(* IEC 61131-3 sources: TetherPLC/tests/tempctrl/cases, 21 files *)

(* ---- t13_handoff.st ---- *)
// t13_handoff.st — the WebUI autotune handoff shape, runtime-verified.
// Mirrors what fbd-lower's expand_st_blocks generates for an inline
// `st` block: VAR_IN_OUT pins aliasing tuner/controller FB instances,
// VAR_OUTPUT live mirrors, and a one-shot APPLY strobe copying gains
// into the controller's input members (CTL.K1 := TUNE.K1 …).
// Same model params as t06 → K1≈6.188 K2≈1.089 Ki≈0.671.
FUNCTION_BLOCK FB_TuneHandoff
VAR_INPUT
    APPLY : BOOL;
    RESET : BOOL;
END_VAR
VAR_OUTPUT
    lqr_k1 : LREAL;
    lqr_k2 : LREAL;
    lqr_ki : LREAL;
    lqr_done : BOOL;
END_VAR
VAR_IN_OUT
    TUNE : FB_AtcLqrTune;
    CTL : FB_AtcLqr;
END_VAR
VAR
    applied : BOOL;
END_VAR
    lqr_k1 := TUNE.K1;
    lqr_k2 := TUNE.K2;
    lqr_ki := TUNE.Ki;
    lqr_done := TUNE.Done;
    IF APPLY AND NOT applied THEN
        CTL.K1 := TUNE.K1;
        CTL.K2 := TUNE.K2;
        CTL.Ki := TUNE.Ki;
        applied := TRUE;
    END_IF;
    IF RESET THEN applied := FALSE; END_IF;
END_FUNCTION_BLOCK

PROGRAM T13
VAR
    flags AT %QB0 : BYTE;
    m : FB_AtcModel2s;
    t : FB_AtcLqrTune;
    c : FB_AtcLqr;
    ho : FB_TuneHandoff;
END_VAR
    m(Execute := TRUE, K := 1.0, Tau := 20.0, Theta := 0.0,
      TauH := 5.0, Ts := 0.5);
    t(Execute := TRUE, A11 := m.A11, A12 := m.A12,
      A21 := m.A21, A22 := m.A22, B1 := m.B1, B2 := m.B2,
      Q1 := 1.0, Q2 := 0.1, Qi := 0.5, R := 1.0, Ts := 0.5,
      MaxIter := 0, Tol := 0.0);
    // K1/K2/Ki intentionally omitted — the handoff owns them; binding
    // them here would clobber the tuned gains every scan (same reason
    // applyTunerToPou strips those params from the controller block).
    c(Execute := FALSE, Setpoint := 0.0, Actual := 0.0,
      X2 := 0.0,
      Nref := 0.0, FFwd := 0.0, OutMin := -100.0, OutMax := 100.0,
      RateLim := 0.0, ManEn := FALSE, ManOut := 0.0,
      CycleTime := 0.1, Reset := FALSE);
    ho(TUNE := t, CTL := c, APPLY := TRUE, RESET := FALSE);
    flags := 0;
    IF t.Done AND t.Conv THEN flags := flags + 1; END_IF;
    IF ABS(ho.lqr_k1 - t.K1) < 0.001 THEN flags := flags + 2; END_IF;
    IF c.K1 > 6.0 AND c.K1 < 6.4 THEN flags := flags + 4; END_IF;
    IF c.K2 > 1.0 AND c.K2 < 1.2 THEN flags := flags + 8; END_IF;
    IF c.Ki > 0.6 AND c.Ki < 0.75 THEN flags := flags + 16; END_IF;
END_PROGRAM

(* ---- t01_math.st ---- *)
// t01_math.st — math function conformance: exp/ln/sqrt/pow against
// known values; flags bit i set when the check passes.
PROGRAM T01
VAR
    flags AT %QB0 : BYTE;
    e1 AT %QD8 : LREAL;
    l1 AT %QD16 : LREAL;
    s1 AT %QD24 : LREAL;
    p1 AT %QD32 : LREAL;
    l2 AT %QD40 : LREAL;
    s2 AT %QD48 : LREAL;
END_VAR
    e1 := F_AtcExp(1.0);          // e = 2.718281828...
    l1 := F_AtcLn(F_AtcExp(3.7)); // = 3.7
    s1 := F_AtcSqrt(2.0);         // 1.41421356...
    p1 := F_AtcPow(2.0, 10.0);    // 1024
    l2 := F_AtcLn(100.0);         // 4.605170186
    s2 := F_AtcSqrt(0.001);       // 0.031622776
    flags := 0;
    IF e1 > 2.718281 AND e1 < 2.718282 THEN flags := flags + 1; END_IF;
    IF l1 > 3.6999 AND l1 < 3.7001 THEN flags := flags + 2; END_IF;
    IF s1 > 1.414213 AND s1 < 1.414214 THEN flags := flags + 4; END_IF;
    IF p1 > 1023.999 AND p1 < 1024.001 THEN flags := flags + 8; END_IF;
    IF l2 > 4.605169 AND l2 < 4.605171 THEN flags := flags + 16; END_IF;
    IF s2 > 0.031622 AND s2 < 0.031624 THEN flags := flags + 32; END_IF;
END_PROGRAM

(* ---- t02_pid.st ---- *)
// t02_pid.st — FB_AtcPid closed loop on a simulated first-order
// plant (K=2 deg/%, Tau=10 s, Ts=0.5 s): PI must pull PV from 20 to
// SP=80 and hold it there. flags: b0 PV in band, b1 output in range,
// b2 Done, b3 no error, b4 anti-windup: output never exceeded 100.
PROGRAM T02
VAR
    flags AT %QB0 : BYTE;
    c : FB_AtcPid;
    pv : LREAL;
    u AT %QD8 : LREAL;
    pvO AT %QD16 : LREAL;
    satHist : LREAL;
END_VAR
    c(Execute := TRUE, Setpoint := 80.0, Actual := pv,
      Kp := 3.0, Tn := 8.0, Tv := 0.0, TfD := 0.0,
      B := 1.0, C := 0.0, FFwd := 0.0,
      OutMin := 0.0, OutMax := 100.0, RateLim := 0.0,
      Deadband := 0.0, HoldI := FALSE, TrackEn := FALSE,
      TrackVal := 0.0, ManEn := FALSE, ManOut := 0.0,
      CycleTime := 0.5, Reset := FALSE);
    u := c.Out;
    IF u > 100.01 OR u < -0.01 THEN
        satHist := 1.0;
    END_IF;
    // plant lag (start PV at 20 deg)
    pv := pv + (2.0 * u - pv) * (0.5 / (10.0 + 0.5));
    pvO := pv;
    flags := 0;
    IF pv > 78.5 AND pv < 82.5 THEN flags := flags + 1; END_IF;
    IF u >= 0.0 AND u <= 100.0 THEN flags := flags + 2; END_IF;
    IF c.Done THEN flags := flags + 4; END_IF;
    IF NOT c.Err THEN flags := flags + 8; END_IF;
    IF satHist = 0.0 THEN flags := flags + 16; END_IF;
END_PROGRAM

(* ---- t03_relay.st ---- *)
// t03_relay.st — FB_AtcRelayTune on a simulated first-order plant
// (K=1, Tau=10 s, Ts=0.5 s): relay hysteresis 2 deg around SP=50,
// MeanOut=50, amp=20. Must finish with Done, plausible Ku/Tu, and
// ZN-classic gains Kp=0.6Ku Tn=0.5Tu Tv=0.125Tu.
// flags: b0 Done, b1 Ku in [4,20], b2 Tu in [4,60], b3 Kp>0,
//        b4 Tn=0.5*Tu, b5 Tv=0.125*Tu, b6 Busy went low, b7 no Err.
PROGRAM T03
VAR
    flags AT %QB0 : BYTE;
    c : FB_AtcRelayTune;
    pv : LREAL;
    u AT %QD8 : LREAL;
    kuO AT %QD16 : LREAL;
    tuO AT %QD24 : LREAL;
END_VAR
    c(Execute := TRUE, Setpoint := 50.0, Actual := pv,
      RelayAmp := 20.0, MeanOut := 50.0, Hyst := 2.0,
      OutMin := 0.0, OutMax := 100.0, TuneRule := 0,
      MinCyc := 3, CycleTime := 0.5,
      Abort := FALSE, Reset := FALSE);
    u := c.Out;
    pv := pv + (1.0 * u - pv) * (0.5 / (10.0 + 0.5));
    kuO := c.Ku;
    tuO := c.Tu;
    flags := 0;
    IF c.Done THEN flags := flags + 1; END_IF;
    IF c.Ku > 4.0 AND c.Ku < 30.0 THEN flags := flags + 2; END_IF;
    IF c.Tu > 4.0 AND c.Tu < 40.0 THEN flags := flags + 4; END_IF;
    IF c.Kp > 0.0 THEN flags := flags + 8; END_IF;
    IF ABS(c.Tn - 0.5 * c.Tu) < 0.01 THEN flags := flags + 16; END_IF;
    IF ABS(c.Tv - 0.125 * c.Tu) < 0.01 THEN flags := flags + 32; END_IF;
    IF NOT c.Busy THEN flags := flags + 64; END_IF;
    IF NOT c.Err THEN flags := flags + 128; END_IF;
END_PROGRAM

(* ---- t04_stepid.st ---- *)
// t04_stepid.st — FB_AtcStepIdent on a simulated FOPDT plant:
// K=2 deg/%, Tau=20 s, true delay 7.5 s (15-scan shift at Ts=0.5),
// step U0=10 -> U1=40. Expect K~2, Tau~20, Theta~7.5+lag bias.
// flags: b0 Done, b1 |K-2|<0.15, b2 14<Tau<28, b3 4<Theta<14,
//        b4 Busy low, b5 no Err, b6 PvFinal ~ K*U1 = 80.
PROGRAM T04
VAR
    flags AT %QB0 : BYTE;
    id : FB_AtcStepIdent;
    pv : LREAL;
    dl : ARRAY[0..15] OF LREAL;
    i : DINT;
    u AT %QD8 : LREAL;
    kO AT %QD16 : LREAL;
    tauO AT %QD24 : LREAL;
    thO AT %QD32 : LREAL;
END_VAR
    id(Execute := TRUE, Actual := pv, U0 := 10.0, U1 := 40.0,
       SettleT := 120.0, TolBand := 0.05, SettleN := 8,
       MaxTime := 600.0, StoreEvery := 4, CycleTime := 0.5,
       Reset := FALSE);
    u := id.Out;
    // plant: 7.5 s transport delay + 20 s lag, gain 2
    pv := pv + (2.0 * dl[15] - pv) * (0.5 / (20.0 + 0.5));
    FOR i := 0 TO 14 DO
        dl[15 - i] := dl[14 - i];
    END_FOR;
    dl[0] := u;
    kO := id.K;
    tauO := id.Tau;
    thO := id.Theta;
    flags := 0;
    IF id.Done THEN flags := flags + 1; END_IF;
    IF id.K > 1.85 AND id.K < 2.15 THEN flags := flags + 2; END_IF;
    IF id.Tau > 14.0 AND id.Tau < 28.0 THEN flags := flags + 4; END_IF;
    IF id.Theta > 4.0 AND id.Theta < 14.0 THEN flags := flags + 8; END_IF;
    IF NOT id.Busy THEN flags := flags + 16; END_IF;
    IF NOT id.Err THEN flags := flags + 32; END_IF;
    IF id.PvFinal > 75.0 AND id.PvFinal < 85.0 THEN
        flags := flags + 64;
    END_IF;
END_PROGRAM

(* ---- t05_rules.st ---- *)
// t05_rules.st — FB_AtcTuneRules on a known FOPDT model
// (K=2, Tau=20, Theta=5). Rule 0 IMC lambda=max(1.25,4)=4:
//   Kp=(20+2.5)/(2*(4+2.5))=1.7308 Tn=22.5 Tv=100/45=2.2222
// Rule 1 SIMC lambda=5: Kp=20/(2*10)=1.0 Tn=min(20,40)=20 Tv=0
// flags: b0 IMC done, b1..3 IMC values, b4 SIMC done, b5 SIMC Kp,
//        b6 ZN done, b7 ZN Kp = 1.2*20/(2*5) = 2.4
PROGRAM T05
VAR
    flags AT %QB0 : BYTE;
    r0 : FB_AtcTuneRules;
    r1 : FB_AtcTuneRules;
    r2 : FB_AtcTuneRules;
    kp0 AT %QD8 : LREAL;
    kp1 AT %QD16 : LREAL;
END_VAR
    r0(Execute := TRUE, K := 2.0, Tau := 20.0, Theta := 5.0,
       Rule := 0, Lambda := 0.0);
    r1(Execute := TRUE, K := 2.0, Tau := 20.0, Theta := 5.0,
       Rule := 1, Lambda := 0.0);
    r2(Execute := TRUE, K := 2.0, Tau := 20.0, Theta := 5.0,
       Rule := 2, Lambda := 0.0);
    kp0 := r0.Kp;
    kp1 := r1.Kp;
    flags := 0;
    IF r0.Done THEN flags := flags + 1; END_IF;
    IF r0.Kp > 1.70 AND r0.Kp < 1.76 THEN flags := flags + 2; END_IF;
    IF r0.Tn > 22.4 AND r0.Tn < 22.6 THEN flags := flags + 4; END_IF;
    IF r0.Tv > 2.2 AND r0.Tv < 2.3 THEN flags := flags + 8; END_IF;
    IF r1.Done THEN flags := flags + 16; END_IF;
    IF r1.Kp > 0.99 AND r1.Kp < 1.01 THEN flags := flags + 32; END_IF;
    IF r2.Done THEN flags := flags + 64; END_IF;
    IF r2.Kp > 2.39 AND r2.Kp < 2.41 THEN flags := flags + 128; END_IF;
END_PROGRAM

(* ---- t06_tuners.st ---- *)
// t06_tuners.st — solvers vs reference values.
// Model from FB_AtcModel2s for K=1 Tau=20 TauH=5 Theta=0 Ts=0.5:
//   a1=e^(-0.025)=0.9753099 a2=e^(-0.1)=0.9048374
//   A=[[.9753,.0247],[0,.9048]] B=[0,0.09516]
// FB_AtcLqrTune Q=diag(1,0.1,0.5) R=1 ->
//   ref (scipy DARE, -Ts aug): K1=6.1884 K2=1.0892 Ki=0.6712
// FB_AtcKalmanTune Q=diag(.01,.01) R=1 -> L1=0.0777 L2=0.00609
// flags: b0/b4 done+conv, b1..3 K in range, b5..6 L in range,
//        b7 model outputs in range
PROGRAM T06
VAR
    flags AT %QB0 : BYTE;
    m : FB_AtcModel2s;
    t : FB_AtcLqrTune;
    kf : FB_AtcKalmanTune;
    k1 AT %QD8 : LREAL;
    k2 AT %QD16 : LREAL;
    ki AT %QD24 : LREAL;
    l1 AT %QD32 : LREAL;
END_VAR
    m(Execute := TRUE, K := 1.0, Tau := 20.0, Theta := 0.0,
      TauH := 5.0, Ts := 0.5);
    t(Execute := TRUE, A11 := m.A11, A12 := m.A12,
      A21 := m.A21, A22 := m.A22, B1 := m.B1, B2 := m.B2,
      Q1 := 1.0, Q2 := 0.1, Qi := 0.5, R := 1.0, Ts := 0.5,
      MaxIter := 0, Tol := 0.0);
    kf(Execute := TRUE, A11 := m.A11, A12 := m.A12,
       A21 := m.A21, A22 := m.A22,
       Q1 := 0.01, Q2 := 0.01, R := 1.0,
       MaxIter := 0, Tol := 0.0);
    k1 := t.K1;
    k2 := t.K2;
    ki := t.Ki;
    l1 := kf.L1;
    flags := 0;
    IF m.Done THEN flags := flags + 1; END_IF;
    IF t.K1 > 6.0 AND t.K1 < 6.4 THEN flags := flags + 2; END_IF;
    IF t.K2 > 1.0 AND t.K2 < 1.2 THEN flags := flags + 4; END_IF;
    IF t.Ki > 0.6 AND t.Ki < 0.75 THEN flags := flags + 8; END_IF;
    IF t.Done AND t.Conv THEN flags := flags + 16; END_IF;
    IF kf.Done AND kf.Conv THEN flags := flags + 32; END_IF;
    IF kf.L1 > 0.07 AND kf.L1 < 0.09 THEN flags := flags + 64; END_IF;
    IF kf.L2 > 0.004 AND kf.L2 < 0.008 THEN flags := flags + 128; END_IF;
END_PROGRAM

(* ---- t07_lqr.st ---- *)
// t07_lqr.st — FB_AtcLqr closed loop on the discrete 2-state sim it
// was tuned for (same A/B as t06). K1=6.1884 K2=1.0892 Ki=0.6712,
// Nref=0 (integral does the tracking). SP=80, x1 starts 0.
// flags: b0 x1 in band, b1 Out in range, b2 Done, b3 no Err,
//        b4 xi finite.
PROGRAM T07
VAR
    flags AT %QB0 : BYTE;
    c : FB_AtcLqr;
    x1 : LREAL;
    x2 : LREAL;
    u AT %QD8 : LREAL;
END_VAR
    c(Execute := TRUE, Setpoint := 80.0, Actual := x1, X2 := x2,
      K1 := 6.1884, K2 := 1.0892, Ki := 0.6712,
      Nref := 0.0, FFwd := 0.0,
      OutMin := 0.0, OutMax := 100.0, RateLim := 0.0,
      ManEn := FALSE, ManOut := 0.0,
      CycleTime := 0.5, Reset := FALSE);
    u := c.Out;
    // plant (discrete, Ts=0.5): x1+ = a1 x1 + (1-a1) x2
    //                         x2+ = a2 x2 + K(1-a2) u
    x1 := 0.9753099 * x1 + 0.0246901 * x2;
    x2 := 0.9048374 * x2 + 0.0951626 * u;
    flags := 0;
    IF x1 > 79.0 AND x1 < 81.0 THEN flags := flags + 1; END_IF;
    IF u >= -0.01 AND u <= 100.01 THEN flags := flags + 2; END_IF;
    IF c.Done THEN flags := flags + 4; END_IF;
    IF NOT c.Err THEN flags := flags + 8; END_IF;
    IF c.Xi > -1.0e6 AND c.Xi < 1.0e6 THEN flags := flags + 16; END_IF;
END_PROGRAM

(* ---- t08_lqg.st ---- *)
// t08_lqg.st — FB_AtcLqg closed loop: same plant as t07 but PV is
// corrupted by a deterministic +/- noise square wave (amplitude 0.5);
// the Kalman filter (L1=0.0777 L2=0.00609) must still track.
// flags: b0 x1 plant state in band, b1 estimated X1 near PV mean,
//        b2 Out bounded, b3 Done, b4 no Err, b5 X2 estimate finite.
PROGRAM T08
VAR
    flags AT %QB0 : BYTE;
    c : FB_AtcLqg;
    x1 : LREAL;
    x2 : LREAL;
    nz : LREAL;
    ymeas : LREAL;
    u AT %QD8 : LREAL;
    xe AT %QD16 : LREAL;
END_VAR
    // deterministic measurement noise: +-0.5 alternating every 7 scans
    nz := nz + 0.5;
    IF nz >= 7.0 THEN nz := -7.0; END_IF;
    ymeas := x1 + nz / 7.0 * 0.5 - 0.25;
    c(Execute := TRUE, Setpoint := 80.0, Actual := ymeas,
      A11 := 0.9753099, A12 := 0.0246901,
      A21 := 0.0, A22 := 0.9048374,
      B1 := 0.0, B2 := 0.0951626,
      L1 := 0.0777, L2 := 0.00609,
      K1 := 6.1884, K2 := 1.0892, Ki := 0.6712,
      Nref := 0.0, FFwd := 0.0,
      OutMin := 0.0, OutMax := 100.0,
      ManEn := FALSE, ManOut := 0.0,
      CycleTime := 0.5, Reset := FALSE);
    u := c.Out;
    x1 := 0.9753099 * x1 + 0.0246901 * x2;
    x2 := 0.9048374 * x2 + 0.0951626 * u;
    xe := c.X1;
    flags := 0;
    IF x1 > 78.0 AND x1 < 82.0 THEN flags := flags + 1; END_IF;
    IF c.X1 > 78.0 AND c.X1 < 82.0 THEN flags := flags + 2; END_IF;
    IF u >= -0.01 AND u <= 100.01 THEN flags := flags + 4; END_IF;
    IF c.Done THEN flags := flags + 8; END_IF;
    IF NOT c.Err THEN flags := flags + 16; END_IF;
    IF c.X2 > -1.0e6 AND c.X2 < 1.0e6 THEN flags := flags + 32; END_IF;
END_PROGRAM

(* ---- t09_profile.st ---- *)
// t09_profile.st — FB_AtcProfile exercising all segment kinds:
//   SEG1 RAMP  -> 100 at 4 deg/s   (PV start 20 -> ~20 s)
//   SEG2 DWELL    100 for 30 s, guaranteed-soak band 2.0
//   SEG3 RAMPT -> 60 in 40 s
//   SEG4 STEP  -> 60 (jump, EV pulse)
//   SEG5 LOOP  -> seg 2, x1 (dwell+rampt run twice)
//   SEG6 END
// Simulated PV lags SP at 10 s. flags: b0 ran to END (Done),
// b1 SP hit 100, b2 SegIdx visited 2, b3 EV word seen (seg2 EV=2),
// b4 guaranteed soak stretched dwell (dwell seg took > 30 s while
// PV lagging outside band... here PV tracks so gsoak rarely bites;
// instead check dwell SegIdx stayed for >= 30 s), b5 loop ran twice
// (saw SegIdx=2 twice => SegIdx reached 4 then 2 again), b6 SP
// finished at 60 (RAMPT target of second pass), b7 no Err.
PROGRAM T09
VAR
    flags AT %QB0 : BYTE;
    prof : FB_AtcProfile;
    pv : LREAL;
    sp AT %QD8 : LREAL;
    segO AT %QD16 : DINT;
    run : BOOL;
    cnt : DINT;
    sawDwell : DINT;
    dwellStart : LREAL;
    dwellLong : BOOL;
    sawSeg4 : BOOL;
    sawLoop : BOOL;
END_VAR
    // ---- segment table (member-wise writes; aggregates can't bind)
    IF cnt = 0 THEN
        prof.SEG[1].KIND := 2;  // RAMP
        prof.SEG[1].TGT := 100.0;
        prof.SEG[1].P1 := 4.0;
        prof.SEG[1].EV := 1;
        prof.SEG[2].KIND := 1;  // DWELL
        prof.SEG[2].TGT := 100.0;
        prof.SEG[2].P1 := 30.0;
        prof.SEG[2].P2 := 2.0;
        prof.SEG[2].EV := 2;
        prof.SEG[3].KIND := 3;  // RAMPT
        prof.SEG[3].TGT := 60.0;
        prof.SEG[3].P1 := 40.0;
        prof.SEG[3].EV := 4;
        prof.SEG[4].KIND := 4;  // STEP
        prof.SEG[4].TGT := 60.0;
        prof.SEG[4].EV := 8;
        prof.SEG[5].KIND := 5;  // LOOP -> seg 2, 1 extra pass
        prof.SEG[5].TGT := 2.0;
        prof.SEG[5].P1 := 1.0;
        prof.SEG[6].KIND := 0;  // END
    END_IF;
    cnt := cnt + 1;
    IF cnt = 2 THEN
        pv := 20.0;   // PV-start point
        run := TRUE;
    END_IF;
    prof(NUM_SEG := 6, RUN := run, HOLD := FALSE, RESET := FALSE,
         PvStart := TRUE, PV := pv, CycleTime := 0.5);
    run := FALSE;
    // simulated PV follows SP (1st-order, 10 s lag)
    pv := pv + (prof.SP - pv) * (0.5 / (10.0 + 0.5));
    sp := prof.SP;
    segO := prof.SegIdx;
    // book-keeping for checks
    IF prof.SegIdx = 2 THEN
        sawDwell := sawDwell + 1;
        IF sawDwell = 1 THEN dwellStart := prof.SegTime; END_IF;
    END_IF;
    IF prof.SegIdx = 2 AND prof.SegTime >= 29.5 THEN
        dwellLong := TRUE;
    END_IF;
    IF prof.SegIdx = 4 THEN sawSeg4 := TRUE; END_IF;
    IF sawSeg4 AND prof.SegIdx = 2 THEN sawLoop := TRUE; END_IF;
    flags := 0;
    IF prof.Done THEN flags := flags + 1; END_IF;
    IF sawDwell >= 2 THEN flags := flags + 2; END_IF;
    IF dwellLong THEN flags := flags + 4; END_IF;
    IF sawSeg4 THEN flags := flags + 8; END_IF;
    IF sawLoop THEN flags := flags + 16; END_IF;
    IF prof.SP > 59.0 AND prof.SP < 61.0 THEN
        flags := flags + 32;
    END_IF;
    IF NOT prof.Err THEN flags := flags + 64; END_IF;
    // extra: the EV word of the END segment is 0; while busy it was
    // nonzero at least once — sawLoop covers seg-2 revisit.
    IF prof.Busy OR prof.Done THEN flags := flags + 128; END_IF;
END_PROGRAM

(* ---- t10_cascade.st ---- *)
// t10_cascade.st — FB_AtcCascadePid: outer product loop (slow, Tau=30)
// drives inner heater loop (fast, Tau=2) setpoint range 20..150;
// inner drives duty 0..100 with gain 1.5 deg/%.
// flags: b0 product PV within band, b1 inner SP clamped to range,
//        b2 Out in range, b3 Done, b4 no Err.
PROGRAM T10
VAR
    flags AT %QB0 : BYTE;
    c : FB_AtcCascadePid;
    pvO : LREAL;
    pvI : LREAL;
    u AT %QD8 : LREAL;
    ispO AT %QD16 : LREAL;
    badIsp : BOOL;
END_VAR
    c(Execute := TRUE, Setpoint := 80.0,
      PvOuter := pvO, PvInner := pvI,
      KpO := 2.0, TnO := 40.0, TvO := 0.0,
      KpI := 4.0, TnI := 4.0, TvI := 0.0,
      InnerSpMin := 20.0, InnerSpMax := 150.0,
      OutMin := 0.0, OutMax := 100.0,
      ManEn := FALSE, ManOut := 0.0,
      CycleTime := 0.5, Reset := FALSE);
    u := c.Out;
    ispO := c.InnerSp;
    IF c.InnerSp < 19.99 OR c.InnerSp > 150.01 THEN
        badIsp := TRUE;
    END_IF;
    // plants: heater lag Tau=2 gain 1.5; product follows heater Tau=30
    pvI := pvI + (1.5 * u - pvI) * (0.5 / (2.0 + 0.5));
    pvO := pvO + (pvI - pvO) * (0.5 / (30.0 + 0.5));
    flags := 0;
    IF pvO > 77.0 AND pvO < 83.0 THEN flags := flags + 1; END_IF;
    IF NOT badIsp THEN flags := flags + 2; END_IF;
    IF u >= -0.01 AND u <= 100.01 THEN flags := flags + 4; END_IF;
    IF c.Done THEN flags := flags + 8; END_IF;
    IF pvI > 0.0 AND pvI <= 150.01 THEN flags := flags + 16; END_IF;
END_PROGRAM

(* ---- t11_smith.st ---- *)
// t11_smith.st — FB_AtcSmith on a dead-time plant:
// K=1 deg/%, Tau=8 s, delay=7.5 s (15 scans); model identical.
// The dead-time compensation must hold SP=60 without oscillation.
// flags: b0 PV in band, b1 Out in range, b2 Done, b3 no Err,
//        b4 model delay state nonzero.
PROGRAM T11
VAR
    flags AT %QB0 : BYTE;
    c : FB_AtcSmith;
    pv : LREAL;
    dl : ARRAY[0..15] OF LREAL;
    i : DINT;
    u AT %QD8 : LREAL;
END_VAR
    c(Execute := TRUE, Setpoint := 60.0, Actual := pv,
      Kp := 0.6, Tn := 10.0, Tv := 0.0,
      ModelK := 1.0, ModelT := 8.0, ModelDt := 7.5,
      OutMin := 0.0, OutMax := 100.0,
      ManEn := FALSE, ManOut := 0.0,
      CycleTime := 0.5, Reset := FALSE);
    u := c.Out;
    // plant: 15-scan delay + 8 s lag, gain 1
    pv := pv + (1.0 * dl[15] - pv) * (0.5 / (8.0 + 0.5));
    FOR i := 0 TO 14 DO
        dl[15 - i] := dl[14 - i];
    END_FOR;
    dl[0] := u;
    flags := 0;
    IF pv > 58.0 AND pv < 62.5 THEN flags := flags + 1; END_IF;
    IF u >= -0.01 AND u <= 100.01 THEN flags := flags + 2; END_IF;
    IF c.Done THEN flags := flags + 4; END_IF;
    IF NOT c.Err THEN flags := flags + 8; END_IF;
    IF c.E > -100.0 AND c.E < 100.0 THEN flags := flags + 16; END_IF;
END_PROGRAM

(* ---- t12_util.st ---- *)
// t12_util.st — signal helpers: FB_AtcPt1, FB_AtcRateLim,
// FB_AtcPwm, FB_AtcHeatCool.
// flags: b0 Pt1 near input after 10*timeconst scans,
//        b1 RateLim respected (|dOut| <= Rate*Ts + eps),
//        b2 Pwm duty ~50% over a period (count on-scans),
//        b3 HeatCool splits (U=-40 -> Cool=40-DeadZone),
//        b4 all Done.
PROGRAM T12
VAR
    flags AT %QB0 : BYTE;
    f1 : FB_AtcPt1;
    rl : FB_AtcRateLim;
    pw : FB_AtcPwm;
    hc : FB_AtcHeatCool;
    cnt : DINT;
    onCnt : DINT;
    pv : LREAL;
    rlPrev : LREAL;
    rlOk : BOOL;
    rlIn : LREAL;
END_VAR
    cnt := cnt + 1;
    // Pt1: step 0->50 at scan 1, Tf=4s
    f1(Execute := TRUE, In := 50.0, Tf := 4.0,
       CycleTime := 0.5, Reset := FALSE);
    pv := f1.Out;
    // RateLim: square wave input +-20, Rate=10/s -> |dOut| <= 5/scan
    IF cnt >= 100 THEN rlIn := -20.0; ELSE rlIn := 20.0; END_IF;
    rl(Execute := TRUE, In := rlIn, Rate := 10.0,
       CycleTime := 0.5, Reset := FALSE);
    IF cnt > 1 THEN
        IF rl.Out - rlPrev > 5.001 OR rl.Out - rlPrev < -5.001 THEN
            rlOk := TRUE;
        END_IF;
    END_IF;
    rlPrev := rl.Out;
    // Pwm: Duty=50, Period=4s (8 scans) — count on-scans over 8 scans
    pw(Execute := TRUE, Duty := 50.0, Period := 4.0, MinOn := 0.0,
       CycleTime := 0.5, Reset := FALSE);
    IF cnt > 190 AND cnt <= 198 THEN
        IF pw.Q THEN onCnt := onCnt + 1; END_IF;
    END_IF;
    // HeatCool: U=-40, dz=2 -> Cool=38*1=38
    hc(Execute := TRUE, U := -40.0, DeadZone := 2.0, CoolGain := 1.0);
    flags := 0;
    IF pv > 48.0 AND pv <= 50.0 THEN flags := flags + 1; END_IF;
    IF NOT rlOk THEN flags := flags + 2; END_IF;
    IF onCnt >= 3 AND onCnt <= 5 THEN flags := flags + 4; END_IF;
    IF hc.Cool > 37.9 AND hc.Cool < 38.1 AND hc.Heat = 0.0 THEN
        flags := flags + 8;
    END_IF;
    IF f1.Done AND rl.Done AND pw.Done AND hc.Done THEN
        flags := flags + 16;
    END_IF;
END_PROGRAM

(* ---- t14_aiscale.st ---- *)
// t14_aiscale.st — FB_AtcAiScale / FB_AtcAoScale: raw int16 channel
// counts <-> engineering units, incl. PT1 filtering and int16
// saturation. Sticky check bits compose into flags %QB0 at the end
// of every scan (idempotent): b0 ai linear exact, b1 ai filtered
// converging, b2 ao roundtrip, b3 ao saturates high, b4 ao
// saturates low -> expect 0x1f.
PROGRAM T14
VAR
    flags AT %QB0 : BYTE;
    ok0, ok1, ok2, ok3, ok4 : BOOL;
    ai : FB_AtcAiScale;
    aoRT : FB_AtcAoScale;
    aoHi : FB_AtcAoScale;
    aoLo : FB_AtcAoScale;
    aiF : FB_AtcAiScale;
    raw : INT;               // analog input channel counts (EL3104-style)
    rawF : INT;              // second channel for the filter test
    counts : INT;            // analog output channel counts (EL4104-style)
    ct : LREAL;
    n : DINT;
END_VAR
    ct := 0.1;
    n := n + 1;

    // ---- AI: EU = Raw*Scale + Offset, no filter
    IF n = 1 THEN raw := 16384; END_IF;
    ai(Execute := TRUE, Raw := raw, Scale := 0.5, Offset := 10.0,
       FiltT := 0.0, CycleTime := ct, Reset := FALSE);
    // 16384 * 0.5 + 10 = 8202
    IF ai.Done AND ai.Out > 8201.9 AND ai.Out < 8202.1 THEN
        ok0 := TRUE;
    END_IF;

    // ---- AI filtered: FiltT=1 s, ct=0.1 -> alpha = 0.1/1.1
    // step rawF 0 -> 1100 counts at n=20; rawf approaches 1100
    IF n = 20 THEN rawF := 1100; END_IF;
    aiF(Execute := TRUE, Raw := rawF, Scale := 1.0, Offset := 0.0,
        FiltT := 1.0, CycleTime := ct, Reset := FALSE);
    // after ~40 filtered steps rawf ~= 1100*(1-(1-alpha)^40) ~ 1080
    IF n >= 40 AND aiF.RawF > 1000.0 AND aiF.RawF < 1100.0 THEN
        ok1 := TRUE;
    END_IF;

    // ---- AO: counts = (In - Offset)/Scale -> int16
    aoRT(Execute := TRUE, In := 8202.0, Scale := 0.5, Offset := 10.0,
         CycleTime := ct, Reset := FALSE);
    IF aoRT.Done AND aoRT.Counts = 16384 AND NOT aoRT.OutBad THEN
        ok2 := TRUE;
    END_IF;

    // ---- AO saturation: way over range -> rail + OutBad
    aoHi(Execute := TRUE, In := 40000.0, Scale := 0.5, Offset := 10.0,
         CycleTime := ct, Reset := FALSE);
    IF aoHi.Done AND aoHi.Counts >= 32767 AND aoHi.OutBad THEN
        ok3 := TRUE;
    END_IF;
    aoLo(Execute := TRUE, In := -40000.0, Scale := 0.5, Offset := 10.0,
         CycleTime := ct, Reset := FALSE);
    IF aoLo.Done AND aoLo.Counts <= -32768 AND aoLo.OutBad THEN
        ok4 := TRUE;
    END_IF;

    flags := 0;
    IF ok0 THEN flags := flags + 1; END_IF;
    IF ok1 THEN flags := flags + 2; END_IF;
    IF ok2 THEN flags := flags + 4; END_IF;
    IF ok3 THEN flags := flags + 8; END_IF;
    IF ok4 THEN flags := flags + 16; END_IF;

    // settle: feed AO counts back to image for observability
    counts := aoRT.Counts;
END_PROGRAM

(* ---- t15_lethality.st ---- *)
// t15_lethality.st — FB_AtcLethality: Tref=70, Z=10, F0Target=1.0 min,
// Temp=90 -> rate=10^2/60=1.667 F0/min, +0.1667/scan. InProduct from
// n=1: F0 hits 1.0 at n=6 (Done). ExitProduct pulse n=4 catches
// acc=0.667<target -> Divert. SensorOK drops n=20 -> Frozen latches;
// ExitProduct n=25 diverts on freeze. Reset n=30 clears acc but the
// same scan re-accumulates, so F0=0.167 at n=30.
// Sticky bits -> flags %QB0: expect 0x3f.
PROGRAM T15
VAR
    flags AT %QB0 : BYTE;
    ok0, ok1, ok2, ok3, ok4, ok5 : BOOL;
    le : FB_AtcLethality;
    n : DINT;
    sok, ex : BOOL;
END_VAR
    n := n + 1;
    sok := NOT (n >= 20 AND n <= 29);
    ex := (n = 4) OR (n = 25);
    le(Temp := 90.0, InProduct := TRUE, SensorOK := sok,
       ExitProduct := ex, Tref := 70.0, Z := 10.0,
       F0Target := 1.0, CycleTime := 0.1,
       Reset := (n = 30));
    IF n = 5 AND le.F0 > 0.5 AND le.F0 < 0.9 THEN ok0 := TRUE; END_IF;
    IF n >= 7 AND n < 15 AND le.Done THEN ok1 := TRUE; END_IF;
    IF n = 4 AND le.Divert THEN ok2 := TRUE; END_IF;
    IF n >= 21 AND n <= 24 AND le.Frozen THEN ok3 := TRUE; END_IF;
    IF n = 25 AND le.Divert THEN ok4 := TRUE; END_IF;
    IF n = 30 AND le.F0 < 0.3 THEN ok5 := TRUE; END_IF;
    flags := 0;
    IF ok0 THEN flags := flags + 1; END_IF;
    IF ok1 THEN flags := flags + 2; END_IF;
    IF ok2 THEN flags := flags + 4; END_IF;
    IF ok3 THEN flags := flags + 8; END_IF;
    IF ok4 THEN flags := flags + 16; END_IF;
    IF ok5 THEN flags := flags + 32; END_IF;
END_PROGRAM

(* ---- t16_heatch.st ---- *)
// t16_heatch.st — FB_AtcHeaterChannel: auto PWM phase, interlock
// inhibit, manual select, and duty clamp. n drives the phases:
//   1-10   auto MV=50%, Period=1s, CycleTime=0.1 -> Q toggles
//   11-20  InterlockOK=FALSE -> Q=FALSE, InterlockBad=TRUE
//   21-30  Auto=FALSE, ManualMV=25 -> DutyApplied=25
//   31-35  MV=150 -> DutyApplied clamped to 100
//   36-45  Execute=FALSE -> Q=FALSE, InterlockBad=FALSE
// Sticky bits -> flags %QB0: expect 0x1f.
PROGRAM T16
VAR
    flags AT %QB0 : BYTE;
    ok0, ok1, ok2, ok3, ok4 : BOOL;
    hc : FB_AtcHeaterChannel;
    n : DINT;
    sawQ : BOOL;
END_VAR
    n := n + 1;
    hc.Execute := n <= 35;
    hc.Enable := TRUE;
    hc.Auto := NOT (n >= 21 AND n <= 30);
    hc.MV := 50.0;
    IF n >= 31 THEN hc.MV := 150.0; END_IF;
    hc.ManualMV := 25.0;
    hc.InterlockOK := NOT (n >= 11 AND n <= 20);
    hc.Period := 1.0;
    hc.MinOn := 0.0;
    hc.CycleTime := 0.1;
    hc();
    IF hc.Q THEN sawQ := TRUE; END_IF;
    ok0 := sawQ;
    IF (n = 15) AND hc.InterlockBad AND NOT hc.Q THEN
        ok1 := TRUE;
    END_IF;
    IF (n = 25) AND (hc.DutyApplied = 25.0) THEN
        ok2 := TRUE;
    END_IF;
    IF (n = 33) AND (hc.DutyApplied = 100.0) THEN
        ok3 := TRUE;
    END_IF;
    IF (n = 40) AND NOT hc.Q AND NOT hc.InterlockBad THEN
        ok4 := TRUE;
    END_IF;
    flags := 0;
    IF ok0 THEN flags := flags + 1; END_IF;
    IF ok1 THEN flags := flags + 2; END_IF;
    IF ok2 THEN flags := flags + 4; END_IF;
    IF ok3 THEN flags := flags + 8; END_IF;
    IF ok4 THEN flags := flags + 16; END_IF;
END_PROGRAM

(* ---- t17_plant.st ---- *)
// t17_plant.st — FB_AtcPlant: FOPDT+deadtime plant simulator.
// Phase 1 (cycles 0..39, U=50 open loop): PV must stay near Pv0
// early (Theta=2 s dead time at 0.5 s scan) then rise toward
// K*U = 100.  Phase 2 (cycles 40+, PI control SP=80): PV settles
// in band.  flags: b0 settled, b1 no err, b2 plant Done,
// b3 output in range, b4 heated above 60, b5 dead time held PV<30
// at cycle 4.
PROGRAM T17
VAR
    flags AT %QB0 : BYTE;
    plant : FB_AtcPlant;
    pid : FB_AtcPid;
    cyc : DINT;
    u : LREAL;
    pvEarly : LREAL;
    maxPv : LREAL;
    closed : BOOL;
END_VAR
    cyc := cyc + 1;
    closed := cyc > 40;
    IF closed THEN
        pid(Execute := TRUE, Setpoint := 80.0, Actual := plant.PV,
            Kp := 3.0, Tn := 8.0, Tv := 0.0, TfD := 0.0,
            B := 1.0, C := 0.0, FFwd := 0.0,
            OutMin := 0.0, OutMax := 100.0, RateLim := 0.0,
            Deadband := 0.0, HoldI := FALSE, TrackEn := FALSE,
            TrackVal := 0.0, ManEn := FALSE, ManOut := 0.0,
            CycleTime := 0.5, Reset := FALSE);
        u := pid.Out;
    ELSE
        u := 50.0;
    END_IF;
    plant(Execute := TRUE, U := u, K := 2.0, Tau1 := 10.0,
          Tau2 := 0.0, Theta := 2.0, Pv0 := 20.0, DistU := 0.0,
          Taamb := 20.0, TauAmb := 0.0, NoiseAmp := 0.0,
          CycleTime := 0.5, Reset := cyc = 1);
    IF cyc = 4 THEN pvEarly := plant.PV; END_IF;
    IF plant.PV > maxPv THEN maxPv := plant.PV; END_IF;
    flags := 0;
    IF closed AND plant.PV > 74.0 AND plant.PV < 86.0 THEN
        flags := flags + 1;
    END_IF;
    IF NOT plant.Err AND NOT pid.Err THEN flags := flags + 2; END_IF;
    IF plant.Done THEN flags := flags + 4; END_IF;
    IF u >= 0.0 AND u <= 100.0 THEN flags := flags + 8; END_IF;
    IF maxPv > 60.0 THEN flags := flags + 16; END_IF;
    IF pvEarly > 0.0 AND pvEarly < 30.0 THEN flags := flags + 32; END_IF;
END_PROGRAM

(* ---- t18_trend.st ---- *)
// t18_trend.st — FB_AtcTrend ring-buffer capture.  Depth=64,
// Value=cycle index, Reset on cycle 1 (records start cycle 2),
// trigger at cycle 20 -> ring pos 18, PostN=4.  72 writes total:
// Wr=70, Full wraps at write 64.
// flags: b0 Done, b1 Full, b2 TrigIdx=18, b3 Buf[TrigIdx]=20
// (trigger sample, not yet overwritten), b4 Count>=40, b5 Wr=72 mod 64 = 8.
PROGRAM T18
VAR
    flags AT %QB0 : BYTE;
    tr : FB_AtcTrend;
    cyc : DINT;
END_VAR
    cyc := cyc + 1;
    tr(Execute := TRUE, CycleTime := 0.1,
       Value := DINT_TO_LREAL(cyc), Depth := 64, PostN := 4,
       Arm := TRUE, Trig := cyc = 20, Reset := cyc = 1);
    flags := 0;
    IF tr.Done THEN flags := flags + 1; END_IF;
    IF tr.Full THEN flags := flags + 2; END_IF;
    IF tr.TrigIdx = 18 THEN flags := flags + 4; END_IF;
    IF tr.TrigIdx >= 0 THEN
        IF tr.Buf[tr.TrigIdx] = 20.0 THEN flags := flags + 8; END_IF;
    END_IF;
    IF tr.Count >= 40 THEN flags := flags + 16; END_IF;
    IF tr.Wr = 8 THEN flags := flags + 32; END_IF;
END_PROGRAM

(* ---- t19_gsched.st ---- *)
// t19_gsched.st — FB_AtcGainSchedule breakpoint interpolation.
// Tables configured once as instance members (array call-args do not
// bind in the MIR), then X varies per call.  X=[0,50,100],
// Kp=[1,2,4], Tn=[10,20,40], Tv=[0,1,2].
// flags: b0 X=0  -> Kp=1 Seg=1 Frac=0
//        b1 X=50 -> Kp=2 Seg=1 Frac=1
//        b2 X=25 -> Kp=1.5 Tn=15 Tv=0.5 Frac=0.5
//        b3 X=75 -> Kp=3 Tn=30 Tv=1.5 Seg=2 Frac=0.5
//        b4 X=-10-> Kp=1 (clamp low)
//        b5 X=200-> Kp=4 (clamp high)
//        b6 dup-X table -> Err
//        b7 X=100-> Kp=4 Seg=2 Frac=1
PROGRAM T19
VAR
    flags AT %QB0 : BYTE;
    gs : FB_AtcGainSchedule;
    gb : FB_AtcGainSchedule;
    cyc : DINT;
END_VAR
    cyc := cyc + 1;
    IF cyc = 1 THEN
        gs.TableX[1] := 0.0;   gs.TableX[2] := 50.0;  gs.TableX[3] := 100.0;
        gs.TableKp[1] := 1.0;  gs.TableKp[2] := 2.0;  gs.TableKp[3] := 4.0;
        gs.TableTn[1] := 10.0; gs.TableTn[2] := 20.0; gs.TableTn[3] := 40.0;
        gs.TableTv[1] := 0.0;  gs.TableTv[2] := 1.0;  gs.TableTv[3] := 2.0;
        gb.TableX := gs.TableX;
        gb.TableKp := gs.TableKp;
        gb.TableTn := gs.TableTn;
        gb.TableTv := gs.TableTv;
        gb.TableX[2] := gb.TableX[1];   // duplicate X -> must flag Err
    END_IF;
    IF cyc >= 2 THEN
        flags := 0;
        gs(Execute := TRUE, X := 0.0, NPts := 3);
        IF gs.Kp = 1.0 AND gs.Seg = 1 AND gs.Frac = 0.0 THEN
            flags := flags + 1;
        END_IF;
        gs(Execute := TRUE, X := 50.0, NPts := 3);
        IF gs.Kp = 2.0 AND gs.Seg = 1 AND gs.Frac = 1.0 THEN
            flags := flags + 2;
        END_IF;
        gs(Execute := TRUE, X := 25.0, NPts := 3);
        IF gs.Kp = 1.5 AND gs.Tn = 15.0 AND gs.Tv = 0.5
           AND gs.Frac = 0.5 THEN
            flags := flags + 4;
        END_IF;
        gs(Execute := TRUE, X := 75.0, NPts := 3);
        IF gs.Kp = 3.0 AND gs.Tn = 30.0 AND gs.Tv = 1.5
           AND gs.Seg = 2 AND gs.Frac = 0.5 THEN
            flags := flags + 8;
        END_IF;
        gs(Execute := TRUE, X := -10.0, NPts := 3);
        IF gs.Kp = 1.0 THEN flags := flags + 16; END_IF;
        gs(Execute := TRUE, X := 200.0, NPts := 3);
        IF gs.Kp = 4.0 THEN flags := flags + 32; END_IF;
        gb(Execute := TRUE, X := 10.0, NPts := 3);
        IF gb.Err THEN flags := flags + 64; END_IF;
        gs(Execute := TRUE, X := 100.0, NPts := 3);
        IF gs.Kp = 4.0 AND gs.Seg = 2 AND gs.Frac = 1.0 THEN
            flags := flags + 128;
        END_IF;
    END_IF;
END_PROGRAM

(* ---- t20_autotune.st ---- *)
// t20_autotune.st — FB_AtcAutoTune end-to-end: relay tune on
// FB_AtcPlant (K=1, Tau=10, Theta=1) drives the plant to a limit
// cycle, gains latch, PID takes over bumplessly via TrackEn.
// flags: b0 at.Done seen, b1 gains sane (Kp>0 Tn>0 Tv>=0 Ku>0 Tu>0),
//        b2 PID settled |PV-50|<10 at end, b3 no Err ever,
//        b4 handoff continuity |dOut|<8 at Done scan,
//        b5 Cycles>=2, b6 PidTrack released after Done,
//        b7 PV stayed in [5,95] whole run.
PROGRAM T20
VAR
    flags AT %QB0 : BYTE;
    aut : FB_AtcAutoTune;
    pid : FB_AtcPid;
    plant : FB_AtcPlant;
    cyc : DINT;
    pvMin : LREAL;
    pvMax : LREAL;
    prevOut : LREAL;
    outAtDone : LREAL;
    dOut : LREAL;
    seenDone : BOOL;
    trackReleased : BOOL;
    inBand : BOOL;
    viol : DINT;
END_VAR
    cyc := cyc + 1;
    IF cyc = 1 THEN
        pvMin := 1.0e9; pvMax := -1.0e9; prevOut := 50.0;
        outAtDone := 0.0; seenDone := FALSE;
        trackReleased := FALSE; inBand := TRUE; viol := 0;
    END_IF;
    aut(Execute := TRUE, Setpoint := 50.0, Actual := plant.PV,
       CycleTime := 0.5, RelayAmp := 20.0, MeanOut := 50.0,
       Hyst := 2.0, OutMin := 0.0, OutMax := 100.0,
       TuneRule := 0, MinCyc := 3, Abort := FALSE, Reset := FALSE,
       PidOut := pid.Out);
    pid(Execute := TRUE, Setpoint := 50.0, Actual := plant.PV,
        Kp := aut.Kp, Tn := aut.Tn, Tv := aut.Tv, TfD := 0.0,
        B := 1.0, C := 0.0, FFwd := 0.0,
        OutMin := 0.0, OutMax := 100.0, RateLim := 0.0,
        Deadband := 0.0, HoldI := FALSE,
        TrackEn := aut.PidTrack, TrackVal := aut.PidTrackVal,
        ManEn := FALSE, ManOut := 0.0,
        CycleTime := 0.5, Reset := cyc = 1);
    plant(Execute := TRUE, U := aut.Out, K := 1.0, Tau1 := 10.0,
          Tau2 := 0.0, Theta := 1.0, Pv0 := 20.0, DistU := 0.0,
          Taamb := 20.0, TauAmb := 0.0, NoiseAmp := 0.0,
          CycleTime := 0.5, Reset := cyc = 1);
    // bookkeeping
    dOut := aut.Out - prevOut;
    IF aut.Done AND NOT seenDone THEN
        seenDone := TRUE;
        outAtDone := aut.Out;
        dOut := aut.Out - prevOut;
    END_IF;
    IF seenDone AND aut.PidTrack = FALSE THEN
        trackReleased := TRUE;
    END_IF;
    IF plant.PV < pvMin THEN pvMin := plant.PV; END_IF;
    IF plant.PV > pvMax THEN pvMax := plant.PV; END_IF;
    IF plant.PV < 5.0 OR plant.PV > 95.0 THEN viol := viol + 1; END_IF;
    IF seenDone AND trackReleased THEN
        IF ABS(plant.PV - 50.0) > 10.0 THEN inBand := FALSE; END_IF;
    END_IF;
    prevOut := aut.Out;
    flags := 0;
    IF aut.Done THEN flags := flags + 1; END_IF;
    IF aut.Kp > 0.0 AND aut.Tn > 0.0 AND aut.Tv >= 0.0
       AND aut.Ku > 0.0 AND aut.Tu > 0.0 THEN
        flags := flags + 2;
    END_IF;
    IF seenDone AND inBand THEN flags := flags + 4; END_IF;
    IF NOT aut.Err THEN flags := flags + 8; END_IF;
    IF seenDone AND ABS(dOut) < 8.0 THEN flags := flags + 16; END_IF;
    IF aut.Cycles >= 2 THEN flags := flags + 32; END_IF;
    IF trackReleased THEN flags := flags + 64; END_IF;
    IF viol = 0 THEN flags := flags + 128; END_IF;
END_PROGRAM

(* ---- t21_recipe.st ---- *)
// t21_recipe.st — FB_AtcBatch: preset-gain profile run with trend.
// 4 segments: RAMP 20->60 @5deg/s (PvStart), DWELL 60 for 20 s,
// RAMP ->30 @5deg/s, END.  PID (preset Kp=3,Tn=12) regulates
// FB_AtcPlant; trend triggers on segment 2.
// flags: b0 Done, b1 Kp stayed preset 3.0, b2 SegIdx hit END (>=4),
//        b3 trend Count>=50, b4 SP reached >=59.5, b5 no Err,
//        b6 trend triggered (TrigIdx>=0), b7 final SP=30.
PROGRAM T21
VAR
    flags AT %QB0 : BYTE;
    rcp : FB_AtcBatch;
    pid : FB_AtcPid;
    plant : FB_AtcPlant;
    cyc : DINT;
    maxSP : LREAL;
    started : BOOL;
END_VAR
    cyc := cyc + 1;
    IF cyc = 1 THEN
        maxSP := 0.0; started := FALSE;
        // segment table (member config, like prof.SEG[i].KIND := ...)
        rcp.SEG[1].KIND := 2;  rcp.SEG[1].TGT := 60.0;
        rcp.SEG[1].P1 := 5.0;  rcp.SEG[1].P2 := 0.0;
        rcp.SEG[2].KIND := 1;  rcp.SEG[2].TGT := 60.0;
        rcp.SEG[2].P1 := 20.0; rcp.SEG[2].P2 := 0.0;
        rcp.SEG[3].KIND := 2;  rcp.SEG[3].TGT := 30.0;
        rcp.SEG[3].P1 := 5.0;  rcp.SEG[3].P2 := 0.0;
        rcp.SEG[4].KIND := 0;
        rcp.nseg := 4;
    END_IF;
    rcp(Execute := TRUE, START := cyc = 2, HOLD := FALSE,
        RESET := cyc = 1, PV := plant.PV, CycleTime := 0.5,
        AutoTune := FALSE, SP_Tune := 50.0,
        RelayAmp := 20.0, MeanOut := 50.0, Hyst := 2.0,
        OutMin := 0.0, OutMax := 100.0, TuneRule := 0, MinCyc := 3,
        AbortTune := FALSE,
        PresetKp := 3.0, PresetTn := 12.0, PresetTv := 0.0,
        TrendEn := TRUE, TrendDepth := 128, PostN := 8,
        TrigSeg := 2, PidOut := pid.Out);
    pid(Execute := TRUE, Setpoint := rcp.SP, Actual := plant.PV,
        Kp := rcp.Kp, Tn := rcp.Tn, Tv := rcp.Tv, TfD := 0.0,
        B := 1.0, C := 0.0, FFwd := 0.0,
        OutMin := 0.0, OutMax := 100.0, RateLim := 0.0,
        Deadband := 0.0, HoldI := FALSE,
        TrackEn := rcp.PidTrack, TrackVal := rcp.PidTrackVal,
        ManEn := FALSE, ManOut := 0.0,
        CycleTime := 0.5, Reset := cyc = 1);
    plant(Execute := TRUE, U := rcp.Out, K := 1.5, Tau1 := 12.0,
          Tau2 := 0.0, Theta := 1.0, Pv0 := 20.0, DistU := 0.0,
          Taamb := 20.0, TauAmb := 0.0, NoiseAmp := 0.0,
          CycleTime := 0.5, Reset := cyc = 1);
    IF rcp.Busy THEN started := TRUE; END_IF;
    IF rcp.SP > maxSP THEN maxSP := rcp.SP; END_IF;
    flags := 0;
    IF rcp.Done THEN flags := flags + 1; END_IF;
    IF rcp.Kp = 3.0 AND rcp.Tn = 12.0 THEN flags := flags + 2; END_IF;
    IF rcp.SegIdx >= 4 THEN flags := flags + 4; END_IF;
    IF rcp.tr.Count >= 50 THEN flags := flags + 8; END_IF;
    IF maxSP >= 59.5 THEN flags := flags + 16; END_IF;
    IF NOT rcp.Err THEN flags := flags + 32; END_IF;
    IF rcp.TrendTrigIdx >= 0 THEN flags := flags + 64; END_IF;
    IF rcp.Done AND rcp.SP = 30.0 THEN flags := flags + 128; END_IF;
END_PROGRAM
